FUNCTION_BLOCK fbShutterCmdSourceHa IMPLEMENTS iShutterCmdSource
VAR_IN_OUT
	HaCmdEvent : stShutterCmdEvent;
END_VAR
VAR
	HaCmdCache : stShutterCmdEvent;
END_VAR

HaCmdCache := HaCmdEvent;

IF HaCmdEvent.Execute THEN
	HaCmdEvent.Execute := FALSE;
END_IF

METHOD Process
VAR_IN_OUT
	CmdEvent	: stShutterCmdEvent;
END_VAR
IF HaCmdCache.Execute THEN
	CmdEvent := HaCmdCache;
	CmdEvent.Source := eShutterCmdSource.HA;
	HaCmdCache.Execute := FALSE;
END_IF
END_METHOD

END_FUNCTION_BLOCK

(* stored: Version 1.1.0.1
   POU fbShutterCmdSourceHa: Id {bea2cbb9-d6f5-424c-a4c2-d3e45d744a98}, SpecialFunc None
   Method Process: Id {577ae5fb-79da-4adc-9275-af801257441c} *)
